Staubli VAL3: pushActCmd.pgx

program pushActCmd(num x_nMoveID, actionIO x_actPrt)
begin
  //add to action stack, excute act command in actCtrl task, to optmize cycle time
  setMutex(bPushToStack)
  _nActStackIndex=(_nActStackIndex+1)%size(actCmd)
  if actCmd[_nActStackIndex].nMoveID<0
    actCmd[_nActStackIndex].nMoveID=x_nMoveID
    actCmd[_nActStackIndex].nActionID =_nActStackIndex
    actPrt[_nActStackIndex]=x_actPrt
  else
    call rs:setAlarm(201,-1)
  endIf
  bPushToStack=false
end
